(* IEC 61131-3 sources: plc-iiot-stack/flagship/tests/POUs/Iiot/FB_IiotKnsMap_Test, 8 files *)

(* ---- FB_IiotKnsMap_Test.decl.st ---- *)
// Назначение: тесты привязки ПЛК-части IIoT-стека к настоящим переменным флагмана КНС-1; выполняются в
//             тестовом приложении флагмана после встраивания (tools_project/flagship_embed.py): значения
//             устройств, станции и регулятора в метриках, инверсия K1, слово тревог станции, запись команд
//             в GVL_Hmi и GVL_Station, счётчик и результат команды станции, PRG_Iiot с подменным клиентом
//             (рождение, метрики тегов флагмана, команда станции до ответа accepted). Глобальные переменные
//             флагмана тест меняет и восстанавливает в том же вызове: другие наборы их не видят.
// Автор:      kr0nsch
// Версия:     0.1.0
// Документ:   docs/TEST_REPORT.md
FUNCTION_BLOCK FB_IiotKnsMap_Test EXTENDS coUnit.FB_TestSuite
VAR
    fbMap : FB_IiotKnsMap;
    aPoints : ARRAY[1..GVL_IiotMap.POINT_COUNT] OF ST_IiotPoint;
    aWords : ARRAY[1..GVL_IiotMap.ALARM_WORDS_COUNT] OF ST_IiotAlarmWords;
    aSmallPoints : ARRAY[1..2] OF ST_IiotPoint;
    aSmallWords : ARRAY[1..2] OF ST_IiotAlarmWords;
END_VAR

(* ---- CmdStateReadsFlagshipCounters.method.decl.st ---- *)
// Счётчик и результат команды: станция — stStationSts, регулятор — fbLIC101.stSts; чужой номер — нули.
METHOD PRIVATE CmdStateReadsFlagshipCounters
VAR
    stStsSaved : ST_StationSts;
    diDev : DINT;
    uiSeq : UINT;
    iResult : INT;
END_VAR

(* ---- CommandsGoToFlagshipCmdStructs.method.decl.st ---- *)
// Принятая команда — в структуру команд флагмана: импульс или значение; строка вне таблицы — FALSE.
METHOD PRIVATE CommandsGoToFlagshipCmdStructs
VAR
    stP102Saved : PL.ST_MotorCmd;
    stP103Saved : PL.ST_MotorCmd;
    stStationSaved : ST_StationCmd;
    stLic101Saved : PL.ST_PidCmd;
    diRule : DINT;
END_VAR

(* ---- FindRule.method.decl.st ---- *)
// Строка белого списка GVL_IiotMap.RULE_CFG для устройства и команды; нет такой — 0.
METHOD PRIVATE FindRule : DINT
VAR_INPUT
    sDevice : STRING(GVL_Const.IIOT_DEVICE_LEN);
    eCommand : E_IiotCommand;
END_VAR
VAR
    diIdx : DINT;
END_VAR

(* ---- FindRule.method.impl.st ---- *)
FindRule := 0;
FOR diIdx := 1 TO GVL_IiotMap.RULE_COUNT DO
    IF GVL_IiotMap.RULE_CFG[diIdx].sDevice = sDevice AND GVL_IiotMap.RULE_CFG[diIdx].eCommand = eCommand THEN
        FindRule := diIdx;
        RETURN;
    END_IF
END_FOR

(* ---- MapReadsFlagshipVariables.method.decl.st ---- *)
// Метрики и слова тревог — из переменных флагмана: K1 инвертируется, режим станции — код перечисления.
METHOD PRIVATE MapReadsFlagshipVariables
VAR
    xK1Saved : BOOL;
    wAlmSaved : WORD;
    eModeSaved : E_StationMode;
END_VAR

(* ---- PrgIiotPublishesAndAppliesStationCommand.method.decl.st ---- *)
// PRG_Iiot с подменным клиентом в приложении флагмана: рождение, метрики тегов флагмана, команда станции
// SetStepped через GVL_Station.stStationCmd до ответа accepted, команда вне белого списка.
METHOD PRIVATE PrgIiotPublishesAndAppliesStationCommand
VAR_INST
    fbFake : FB_MqttClientFake;
    xRan : BOOL;              // тест длинный: выполняется один раз, дальше coUnit только вызывает метод
END_VAR
VAR
    iCall : INT;
    uliNow : ULINT;
    stCmdSaved : ST_StationCmd;
    stStsSaved : ST_StationSts;
    xK1Saved : BOOL;
    sCmd : STRING(GVL_Const.MQTT_CMD_PAYLOAD_LEN);
END_VAR

(* ---- PrgIiotPublishesAndAppliesStationCommand.method.impl.st ---- *)
coUnit.TEST('PrgIiotPublishesAndAppliesStationCommand');

IF xRan THEN
    coUnit.TEST_FINISHED();
    RETURN;
END_IF
xRan := TRUE;
stCmdSaved := GVL_Station.stStationCmd;
stStsSaved := GVL_Station.stStationSts;
xK1Saved := GVL_IO.xK1;
fbFake.aCapture[1] := 'vodokanal/kns1/station/PLC1/status/connection';
fbFake.aCapture[2] := 'vodokanal/kns1/station/K1/general_alarm';
fbFake.aCapture[3] := 'vodokanal/kns1/station/KNS1/mode';
fbFake.aCapture[4] := 'vodokanal/kns1/station/LIC101/pv';
fbFake.aCapture[5] := 'vodokanal/kns1/station/KNS1/cmd_ack/SetStepped';
fbFake.aCapture[6] := 'vodokanal/kns1/station/V1/cmd_ack/SetOos';
GVL_IO.xK1 := FALSE;
GVL_Station.stStationSts.eMode := E_StationMode.Auto;
GVL_Iiot.stIiotCfg.xEnable := TRUE;
GVL_Iiot.stIiotCfg.xCommandsEnable := TRUE;
PRG_Iiot.itfClientOverride := fbFake;
FOR iCall := 1 TO 60 DO   // 139 метрик по 8 и 88 тревог по 4 за цикл, с запасом
    PRG_Iiot();
END_FOR
AssertTrue(Condition := GVL_Iiot.stIiotSts.eConnState = E_MqttConnState.Connected AND GVL_Iiot.stIiotSts.xClockValid,
           Message := 'connected with a valid clock');
AssertTrue(Condition := fbFake.LastHas(sTopic := 'vodokanal/kns1/station/PLC1/status/connection',
           sPart := '"node":"PLC1","state":"online","reason":"birth","source":"codesys"'), Message := 'birth');
AssertTrue(Condition := fbFake.LastHas(sTopic := 'vodokanal/kns1/station/K1/general_alarm', sPart := '"value":1,'),
           Message := CONCAT('K1 released -> 1: ',
                             fbFake.LastPayload(sTopic := 'vodokanal/kns1/station/K1/general_alarm')));
AssertTrue(Condition := fbFake.LastHas(sTopic := 'vodokanal/kns1/station/KNS1/mode', sPart := '"value":1,'),
           Message := CONCAT('station mode Auto -> 1: ',
                             fbFake.LastPayload(sTopic := 'vodokanal/kns1/station/KNS1/mode')));
AssertEquals_UINT(Expected := 1, Actual := fbFake.CountTopic(sTopic := 'vodokanal/kns1/station/LIC101/pv'),
                  Message := 'LIC101 pv published once');
AssertEquals_UINT(Expected := 0, Actual := GVL_Iiot.stIiotSts.uiQueue, Message := 'everything published');

// команда станции SetStepped: шлюз -> GVL_Station.stStationCmd -> обработка станцией -> ответ accepted
SysTimeRtcHighResGet(pTimestamp := uliNow);
sCmd := CONCAT(CONCAT('{"schema_version":"1.1","cmd_id":"kns00001","ts":', ULINT_TO_STRING(uliNow)),
               ',"origin":"test","command":"SetStepped"}');
GVL_Station.stStationCmd.xSetStepped := FALSE;
fbFake.Inject(sTopic := 'vodokanal/kns1/station/KNS1/cmd/SetStepped', sPayload := sCmd, xTruncated := FALSE,
              xRetained := FALSE);
PRG_Iiot();
AssertTrue(Condition := GVL_Station.stStationCmd.xSetStepped,
           Message := 'SetStepped -> GVL_Station.stStationCmd.xSetStepped');
AssertEquals_UINT(Expected := 0,
                  Actual := fbFake.CountTopic(sTopic := 'vodokanal/kns1/station/KNS1/cmd_ack/SetStepped'),
                  Message := 'no ack before the station processed the command');
// станция обработала команду (в тестовом приложении PRG_Station не вызывается — её ответ пишет тест)
GVL_Station.stStationSts.uiCmdSeq := GVL_Station.stStationSts.uiCmdSeq + 1;
GVL_Station.stStationSts.eCmdResult := PL.E_CmdResult.Accepted;
PRG_Iiot();
AssertTrue(Condition := fbFake.LastHas(sTopic := 'vodokanal/kns1/station/KNS1/cmd_ack/SetStepped',
           sPart := '"cmd_id":"kns00001"'), Message := 'ack for kns00001');
AssertTrue(Condition := fbFake.LastHas(sTopic := 'vodokanal/kns1/station/KNS1/cmd_ack/SetStepped',
           sPart := '"result":"accepted","reason":"ok"}'),
           Message := CONCAT('accepted after the station processed the command: ',
                             fbFake.LastPayload(sTopic := 'vodokanal/kns1/station/KNS1/cmd_ack/SetStepped')));
// SetOos не в белом списке
sCmd := CONCAT(CONCAT('{"schema_version":"1.1","cmd_id":"kns00002","ts":', ULINT_TO_STRING(uliNow)),
               ',"origin":"test","command":"SetOos"}');
fbFake.Inject(sTopic := 'vodokanal/kns1/station/V1/cmd/SetOos', sPayload := sCmd, xTruncated := FALSE,
              xRetained := FALSE);
PRG_Iiot();
AssertTrue(Condition := fbFake.LastHas(sTopic := 'vodokanal/kns1/station/V1/cmd_ack/SetOos',
           sPart := '"result":"rejected","reason":"not_whitelisted"}'), Message := 'SetOos rejected');
AssertEquals_UDINT(Expected := 1, Actual := GVL_Iiot.stIiotSts.udiCmdAccepted, Message := 'one accepted');

// обмен выключен: штатное отключение; глобальные переменные флагмана — как были
GVL_Iiot.stIiotCfg.xEnable := FALSE;
GVL_Iiot.stIiotCfg.xCommandsEnable := FALSE;
PRG_Iiot();
AssertTrue(Condition := fbFake.LastHas(sTopic := 'vodokanal/kns1/station/PLC1/status/connection',
           sPart := '"state":"offline","reason":"shutdown"'), Message := 'shutdown status');
PRG_Iiot.itfClientOverride := 0;
PRG_Iiot();
GVL_Station.stStationCmd := stCmdSaved;
GVL_Station.stStationSts := stStsSaved;
GVL_IO.xK1 := xK1Saved;

coUnit.TEST_FINISHED();
